FUNCTION_BLOCK ButtonsPanel (* Composite Function Block Type *)
  (* Standard: 61499-2 *)
  (* Version 0.0, 7/13/2016, Andrei, nxtControl GmbH, template *)
  PACKAGE Main;
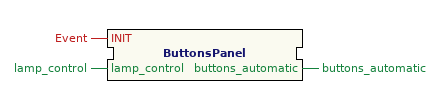
  EVENT_INPUT
    INIT; (* Initialization Request *)
  END_EVENT
  SOCKETS
    lamp_control : lamp_control;
  END_SOCKETS
  PLUGS
    buttons_automatic : buttons_automatic;
  END_PLUGS
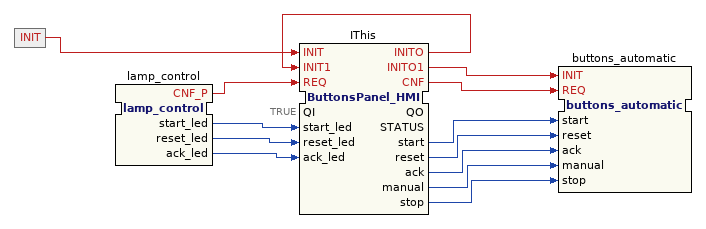
  FBS
    IThis : ButtonsPanel_HMI(QI := TRUE);
  END_FBS
  EVENT_CONNECTIONS
    INIT TO IThis.INIT;
    IThis.INITO TO IThis.INIT1;
    lamp_control.CNF_P TO IThis.REQ;
    IThis.INITO1 TO buttons_automatic.INIT;
    IThis.CNF TO buttons_automatic.REQ;
  END_CONNECTIONS
  DATA_CONNECTIONS
    lamp_control.start_led TO IThis.start_led;
    lamp_control.reset_led TO IThis.reset_led;
    lamp_control.ack_led TO IThis.ack_led;
    IThis.start TO buttons_automatic.start;
    IThis.reset TO buttons_automatic.reset;
    IThis.ack TO buttons_automatic.ack;
    IThis.manual TO buttons_automatic.manual;
    IThis.stop TO buttons_automatic.stop;
  END_CONNECTIONS
END_FUNCTION_BLOCK
